FUNCTION_BLOCK basicAguaReuso (* Logica unica da agua de reuso (PIT-01/02, boia LSL-01, comunicacao) *)
  (* Standard: 61499-2 *)
  (* Version 1.2, 15/10/2026, Hidryco, Hidryco, 1.2: sai o MGE (vira instancia propria no ETE_TJ). 1.0: monitoracao da agua de reuso - niveis 1000-PIT-01/02, boia 1000-LSL-01 e comunicacao das remotas 1/2 da Subestacao *)
  PACKAGE Hidryco.HidrycoLib;
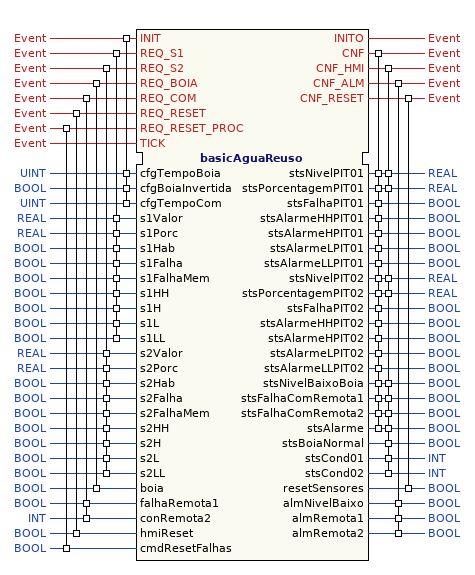
  EVENT_INPUT
    INIT WITH cfgTempoBoia, cfgBoiaInvertida, cfgTempoCom; (* Inicializacao *)
    REQ_S1 WITH s1Valor, s1Porc, s1Hab, s1Falha, s1FalhaMem, s1HH, s1H, s1L, s1LL; (* PIT_1000_01 *)
    REQ_S2 WITH s2Valor, s2Porc, s2Hab, s2Falha, s2FalhaMem, s2HH, s2H, s2L, s2LL; (* PIT_1000_02 *)
    REQ_BOIA WITH boia; (* Boia 1000-LSL-01 *)
    REQ_COM WITH falhaRemota1, conRemota2; (* Comunicacao das remotas *)
    REQ_RESET WITH hmiReset; (* Reset pela IHM *)
    REQ_RESET_PROC WITH cmdResetFalhas; (* Reset pelo processo *)
    TICK; (* Base de tempo de 1 s (E_CYCLE) *)
  END_EVENT
  EVENT_OUTPUT
    INITO; (* Inicializacao concluida *)
    CNF WITH stsNivelPIT01, stsPorcentagemPIT01, stsFalhaPIT01, stsAlarmeHHPIT01, stsAlarmeHPIT01, stsAlarmeLPIT01, stsAlarmeLLPIT01, stsNivelPIT02, stsPorcentagemPIT02, stsFalhaPIT02, stsAlarmeHHPIT02, stsAlarmeHPIT02, stsAlarmeLPIT02, stsAlarmeLLPIT02, stsNivelBaixoBoia, stsFalhaComRemota1, stsFalhaComRemota2, stsAlarme; (* Valores e alarmes para o processo (na mudanca) *)
    CNF_HMI WITH stsNivelPIT01, stsPorcentagemPIT01, stsNivelPIT02, stsPorcentagemPIT02, stsCond01, stsCond02, stsBoiaNormal, stsNivelBaixoBoia, stsFalhaComRemota1, stsFalhaComRemota2, stsAlarme; (* Status para a IHM (na mudanca) *)
    CNF_ALM WITH almNivelBaixo, almRemota1, almRemota2; (* Alarmes para os ALARM_BIT (na mudanca) *)
    CNF_RESET WITH resetSensores; (* Reset dos sensores *)
  END_EVENT
  VAR_INPUT
    cfgTempoBoia : UINT := 10; (* Tempo (s) da boia 1000-LSL-01 abaixada para confirmar o nivel baixo *)
    cfgBoiaInvertida : BOOL := FALSE; (* FALSE: entrada da boia TRUE = nivel normal (boia levantada). TRUE: entrada TRUE = nivel baixo *)
    cfgTempoCom : UINT := 5; (* Tempo (s) sem comunicacao para confirmar a falha das remotas *)
    s1Valor : REAL; (* PIT_1000_01: valor (stsValor) *)
    s1Porc : REAL; (* PIT_1000_01: porcentagem (stsPorcentagem) *)
    s1Hab : BOOL; (* PIT_1000_01: sensor habilitado *)
    s1Falha : BOOL; (* PIT_1000_01: sinal invalido agora (stsFalhaAtiva) *)
    s1FalhaMem : BOOL; (* PIT_1000_01: falha do sensor memorizada (stsFalhaSensor) *)
    s1HH : BOOL; (* PIT_1000_01: alarme HH *)
    s1H : BOOL; (* PIT_1000_01: alarme H *)
    s1L : BOOL; (* PIT_1000_01: alarme L *)
    s1LL : BOOL; (* PIT_1000_01: alarme LL *)
    s2Valor : REAL; (* PIT_1000_02: valor (stsValor) *)
    s2Porc : REAL; (* PIT_1000_02: porcentagem (stsPorcentagem) *)
    s2Hab : BOOL; (* PIT_1000_02: sensor habilitado *)
    s2Falha : BOOL; (* PIT_1000_02: sinal invalido agora (stsFalhaAtiva) *)
    s2FalhaMem : BOOL; (* PIT_1000_02: falha do sensor memorizada (stsFalhaSensor) *)
    s2HH : BOOL; (* PIT_1000_02: alarme HH *)
    s2H : BOOL; (* PIT_1000_02: alarme H *)
    s2L : BOOL; (* PIT_1000_02: alarme L *)
    s2LL : BOOL; (* PIT_1000_02: alarme LL *)
    boia : BOOL; (* Campo: boia 1000-LSL-01 (remota 1 da Subestacao, A6 %I0.105) *)
    falhaRemota1 : BOOL; (* Campo: falha de comunicacao da remota 1 da Subestacao (FALHA_COM do cartao SUB_R1_A6_DI32K0) *)
    conRemota2 : INT; (* Campo: connStatusInt da remota 2 da Subestacao (1 = online) *)
    hmiReset : BOOL; (* IHM: reset / reconhecimento *)
    cmdResetFalhas : BOOL; (* Processo: reset (com E_RESET_FALHAS) *)
  END_VAR
  VAR_OUTPUT
    stsNivelPIT01 : REAL; (* Nivel PIT_1000_01 (unidade de engenharia do sensor; 0 com o sinal em falha) *)
    stsPorcentagemPIT01 : REAL; (* Nivel PIT_1000_01 em % da altura maxima *)
    stsFalhaPIT01 : BOOL; (* Falha do sensor PIT_1000_01 (memorizada ate o reset) *)
    stsAlarmeHHPIT01 : BOOL; (* Alarme HH do PIT_1000_01 *)
    stsAlarmeHPIT01 : BOOL; (* Alarme H do PIT_1000_01 *)
    stsAlarmeLPIT01 : BOOL; (* Alarme L do PIT_1000_01 *)
    stsAlarmeLLPIT01 : BOOL; (* Alarme LL do PIT_1000_01 *)
    stsNivelPIT02 : REAL; (* Nivel PIT_1000_02 (unidade de engenharia do sensor; 0 com o sinal em falha) *)
    stsPorcentagemPIT02 : REAL; (* Nivel PIT_1000_02 em % da altura maxima *)
    stsFalhaPIT02 : BOOL; (* Falha do sensor PIT_1000_02 (memorizada ate o reset) *)
    stsAlarmeHHPIT02 : BOOL; (* Alarme HH do PIT_1000_02 *)
    stsAlarmeHPIT02 : BOOL; (* Alarme H do PIT_1000_02 *)
    stsAlarmeLPIT02 : BOOL; (* Alarme L do PIT_1000_02 *)
    stsAlarmeLLPIT02 : BOOL; (* Alarme LL do PIT_1000_02 *)
    stsNivelBaixoBoia : BOOL; (* Nivel baixo pela boia 1000-LSL-01 (confirmado por cfgTempoBoia) *)
    stsFalhaComRemota1 : BOOL; (* Falha de comunicacao com a remota 1 da Subestacao (boia) *)
    stsFalhaComRemota2 : BOOL; (* Falha de comunicacao com a remota 2 da Subestacao (PIT-01/02) *)
    stsAlarme : BOOL; (* Algum alarme da agua de reuso (sensores, boia, comunicacao) *)
    stsBoiaNormal : BOOL; (* Boia 1000-LSL-01 levantada (nivel acima do baixo) *)
    stsCond01 : INT; (* PIT-01 para a IHM: 0 normal, 1 HH, 2 H, 3 L, 4 LL, 5 sinal invalido, 6 falha memorizada, 7 desabilitado *)
    stsCond02 : INT; (* PIT-02 para a IHM (mesmos codigos) *)
    resetSensores : BOOL; (* Reset dos sensores (com CNF_RESET) *)
    almNivelBaixo : BOOL; (* ALARM_BIT nivel baixo (boia) *)
    almRemota1 : BOOL; (* ALARM_BIT remota 1 *)
    almRemota2 : BOOL; (* ALARM_BIT remota 2 *)
  END_VAR
  VAR
    initDone : BOOL;
    initPass : BOOL;
    bReset : BOOL;
    bBoiaRecebida : BOOL; (* Ja houve leitura da boia *)
    bCondBaixo : BOOL; (* Boia abaixada agora (remota 1 ok) *)
    uSegBoia : UDINT;
    uSegRem1 : UDINT;
    uSegRem2 : UDINT;
    bRem2 : BOOL;
    wSts : WORD;
    oldSts : WORD := 16#FFFF;
    wAlm : WORD;
    oldAlm : WORD := 16#FFFF;
    oldN1 : REAL := -1.0;
    oldP1 : REAL := -1.0;
    oldN2 : REAL := -1.0;
    oldP2 : REAL := -1.0;
    oldC1 : INT := -1;
    oldC2 : INT := -1;
  END_VAR
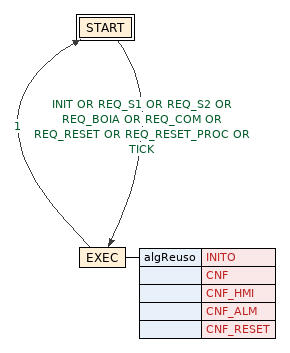
  EC_STATES
    START; (* Estado inicial *)
    EXEC : algReuso -> INITO, -> CNF, -> CNF_HMI, -> CNF_ALM, -> CNF_RESET; (* Executa a logica; o algoritmo decide quais eventos saem *)
  END_STATES
  EC_TRANSITIONS
    START TO EXEC := INIT OR REQ_S1 OR REQ_S2 OR REQ_BOIA OR REQ_COM OR REQ_RESET OR REQ_RESET_PROC OR TICK;
    EXEC TO START := 1;
  END_TRANSITIONS
  ALGORITHM algReuso IN ST: (* Logica completa da agua de reuso (um unico algoritmo) *)
(* =====================================================================
   basicAguaReuso v1.2 - Agua de reuso (serie 1000) - so monitoracao
   Padrao das bibliotecas Schneider: eventos de saida desligados no inicio e
   ligados so na mudanca; tempos contados pelo TICK de 1 s (E_CYCLE do CAT).
   - 1000-PIT-01 / 1000-PIT-02: Sensor_Generico (4-20 mA, nivel); valores,
     falha e alarmes HH/H/L/LL repassados para as saidas do CAT;
   - boia 1000-LSL-01: nivel baixo depois de cfgTempoBoia s abaixada;
     ignorada com a remota 1 em falha (os bits ficam congelados);
   - falha de comunicacao: remota 1 (cartao) e remota 2 (connStatusInt
     diferente de 1) confirmada depois de cfgTempoCom s;
   - v1.2: o MGE do PCM Agua Reuso saiu daqui: e a instancia MGE_AGUA_REUSO
     (MGE_Generico) no frame dos MGEs do layer ETE_TJ;
   - reset (IHM ou processo): reset dos sensores; a IHM tambem reconhece.
   ===================================================================== *)

(* ---- 0. Eventos de saida: so sai o que for ligado abaixo ---- *)
INITO     := FALSE;
CNF       := FALSE;
CNF_HMI   := FALSE;
CNF_ALM   := FALSE;
CNF_RESET := FALSE;

IF REQ_BOIA THEN
    bBoiaRecebida := TRUE;
END_IF;

(* ---- 1. Inicializacao ---- *)
IF INIT THEN
    initDone := TRUE;
    initPass := TRUE;
    INITO    := TRUE;
END_IF;
IF NOT initDone THEN
    RETURN;
END_IF;

(* ---- 2. Reset ---- *)
bReset := (REQ_RESET AND hmiReset) OR (REQ_RESET_PROC AND cmdResetFalhas);
IF bReset THEN
    resetSensores := TRUE;
    CNF_RESET := TRUE;
END_IF;

(* ---- 3. Comunicacao (falha confirmada depois de cfgTempoCom s) ---- *)
IF falhaRemota1 THEN
    IF TICK AND uSegRem1 < UINT_TO_UDINT(cfgTempoCom) THEN
        uSegRem1 := uSegRem1 + 1;
    END_IF;
ELSE
    uSegRem1 := 0;
END_IF;
stsFalhaComRemota1 := falhaRemota1 AND uSegRem1 >= UINT_TO_UDINT(cfgTempoCom);

bRem2 := conRemota2 <> 1;
IF bRem2 THEN
    IF TICK AND uSegRem2 < UINT_TO_UDINT(cfgTempoCom) THEN
        uSegRem2 := uSegRem2 + 1;
    END_IF;
ELSE
    uSegRem2 := 0;
END_IF;
stsFalhaComRemota2 := bRem2 AND uSegRem2 >= UINT_TO_UDINT(cfgTempoCom);

(* ---- 4. Boia 1000-LSL-01 ---- *)
stsBoiaNormal := boia XOR cfgBoiaInvertida;      (* TRUE = boia levantada (nivel acima do baixo) *)
bCondBaixo := bBoiaRecebida AND NOT falhaRemota1 AND NOT stsBoiaNormal;
IF bCondBaixo THEN
    IF TICK AND uSegBoia < UINT_TO_UDINT(cfgTempoBoia) THEN
        uSegBoia := uSegBoia + 1;
    END_IF;
ELSE
    uSegBoia := 0;
END_IF;
stsNivelBaixoBoia := bCondBaixo AND uSegBoia >= UINT_TO_UDINT(cfgTempoBoia);

(* ---- 5. Sensores ---- *)
stsNivelPIT01 := s1Valor;
stsPorcentagemPIT01 := s1Porc;
stsFalhaPIT01 := s1FalhaMem;
stsAlarmeHHPIT01 := s1HH;
stsAlarmeHPIT01 := s1H;
stsAlarmeLPIT01 := s1L;
stsAlarmeLLPIT01 := s1LL;
stsNivelPIT02 := s2Valor;
stsPorcentagemPIT02 := s2Porc;
stsFalhaPIT02 := s2FalhaMem;
stsAlarmeHHPIT02 := s2HH;
stsAlarmeHPIT02 := s2H;
stsAlarmeLPIT02 := s2L;
stsAlarmeLLPIT02 := s2LL;

(* condicao para a IHM, da mais grave para a menos grave *)
IF NOT s1Hab THEN
    stsCond01 := 7;
ELSIF s1Falha THEN
    stsCond01 := 5;
ELSIF s1FalhaMem THEN
    stsCond01 := 6;
ELSIF s1HH THEN
    stsCond01 := 1;
ELSIF s1LL THEN
    stsCond01 := 4;
ELSIF s1H THEN
    stsCond01 := 2;
ELSIF s1L THEN
    stsCond01 := 3;
ELSE
    stsCond01 := 0;
END_IF;
IF NOT s2Hab THEN
    stsCond02 := 7;
ELSIF s2Falha THEN
    stsCond02 := 5;
ELSIF s2FalhaMem THEN
    stsCond02 := 6;
ELSIF s2HH THEN
    stsCond02 := 1;
ELSIF s2LL THEN
    stsCond02 := 4;
ELSIF s2H THEN
    stsCond02 := 2;
ELSIF s2L THEN
    stsCond02 := 3;
ELSE
    stsCond02 := 0;
END_IF;

(* ---- 6. Alarmes ---- *)
almNivelBaixo := stsNivelBaixoBoia;
almRemota1 := stsFalhaComRemota1;
almRemota2 := stsFalhaComRemota2;
stsAlarme := s1FalhaMem OR s1HH OR s1H OR s1L OR s1LL OR s2FalhaMem OR s2HH OR s2H OR s2L OR s2LL
             OR almNivelBaixo OR almRemota1 OR almRemota2;

(* ---- 7. Eventos so na mudanca ---- *)
wSts := 0;
IF stsFalhaPIT01      THEN wSts := wSts OR 16#0001; END_IF;
IF stsAlarmeHHPIT01   THEN wSts := wSts OR 16#0002; END_IF;
IF stsAlarmeHPIT01    THEN wSts := wSts OR 16#0004; END_IF;
IF stsAlarmeLPIT01    THEN wSts := wSts OR 16#0008; END_IF;
IF stsAlarmeLLPIT01   THEN wSts := wSts OR 16#0010; END_IF;
IF stsFalhaPIT02      THEN wSts := wSts OR 16#0020; END_IF;
IF stsAlarmeHHPIT02   THEN wSts := wSts OR 16#0040; END_IF;
IF stsAlarmeHPIT02    THEN wSts := wSts OR 16#0080; END_IF;
IF stsAlarmeLPIT02    THEN wSts := wSts OR 16#0100; END_IF;
IF stsAlarmeLLPIT02   THEN wSts := wSts OR 16#0200; END_IF;
IF stsNivelBaixoBoia  THEN wSts := wSts OR 16#0400; END_IF;
IF stsFalhaComRemota1 THEN wSts := wSts OR 16#0800; END_IF;
IF stsFalhaComRemota2 THEN wSts := wSts OR 16#1000; END_IF;
IF stsAlarme          THEN wSts := wSts OR 16#4000; END_IF;
IF stsBoiaNormal      THEN wSts := wSts OR 16#8000; END_IF;
CNF := initPass OR ((wSts AND 16#7FFF) <> (oldSts AND 16#7FFF)) OR (stsNivelPIT01 <> oldN1) OR (stsPorcentagemPIT01 <> oldP1)
       OR (stsNivelPIT02 <> oldN2) OR (stsPorcentagemPIT02 <> oldP2);
CNF_HMI := initPass OR (wSts <> oldSts) OR (stsNivelPIT01 <> oldN1) OR (stsPorcentagemPIT01 <> oldP1)
           OR (stsNivelPIT02 <> oldN2) OR (stsPorcentagemPIT02 <> oldP2) OR (stsCond01 <> oldC1) OR (stsCond02 <> oldC2);
wAlm := 0;
IF almNivelBaixo THEN wAlm := wAlm OR 16#0001; END_IF;
IF almRemota1    THEN wAlm := wAlm OR 16#0002; END_IF;
IF almRemota2    THEN wAlm := wAlm OR 16#0004; END_IF;
CNF_ALM := initPass OR (wAlm <> oldAlm);
oldSts := wSts;
oldAlm := wAlm;
oldN1 := stsNivelPIT01;
oldP1 := stsPorcentagemPIT01;
oldN2 := stsNivelPIT02;
oldP2 := stsPorcentagemPIT02;
oldC1 := stsCond01;
oldC2 := stsCond02;

initPass := FALSE;
  END_ALGORITHM
END_FUNCTION_BLOCK
